(* CODESYS project Diagnosis.vis.xml

Project tree, tasks and I/O mapping:
  visualisation Diagnosis
*)

// /Diagnosis
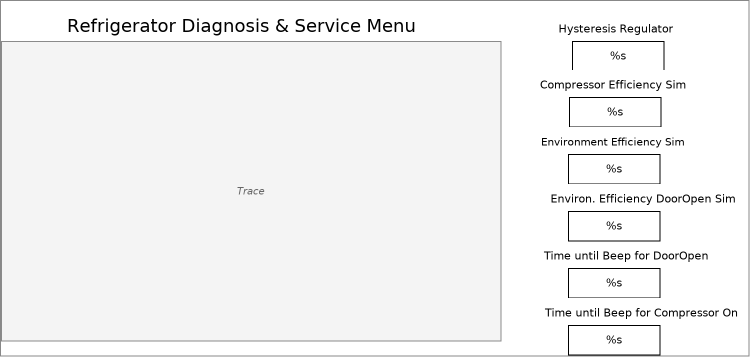
VISUALIZATION Diagnosis  // 750x357
    Trace (1,41 500x300)
    Rectangle (24,11 435x30), "Refrigerator Diagnosis & Service Menu"
    Group (541,14 150x57)
        Rectangle (0,0 150x30), "Hysteresis Regulator"
        Rectangle (31,27 92x30), "%s", text variable: PLC_PRG.Hysteresis
            OnMouseDown: write the text variable via Default
    Group (538,70 150x57)
        Rectangle (0,0 150x30), "Compressor Efficiency Sim"
        Rectangle (31,27 92x30), "%s", text variable: Simulation.P_Cooling
            OnMouseDown: write the text variable via Default
    Group (538,127 150x57)
        Rectangle (0,0 150x30), "Environment Efficiency Sim"
        Rectangle (30,27 92x30), "%s", text variable: Simulation.P_Environment
            OnMouseDown: write the text variable via Default
    Group (538,241 177x57)
        Rectangle (0,0 177x30), "Time until Beep for DoorOpen"
        Rectangle (30,27 92x30), "%s", text variable: Glob_Var.DoorOpenThreshold
            OnMouseDown: write the text variable via Default
    Group (538,298 207x57)
        Rectangle (0,0 207x30), "Time until Beep for Compressor On"
        Rectangle (30,27 92x30), "%s", text variable: Glob_Var.AlarmThreshold
            OnMouseDown: write the text variable via Default
    Rectangle (538,184 210x30), "Environ. Efficiency DoorOpen Sim"
    Rectangle (568,211 92x30), "%s", text variable: Simulation.P_EnvironmentDoorOpen
        OnMouseDown: write the text variable via Default
END_VISUALIZATION
